Universal Robots PolyScope program: TgtProg.urp

Program TgtProg (createdIn=3.0.0 lastSavedIn=3.0.0 directory=/programs installation=default)
Robot Program (runOnlyOnce=true motionType=MoveJ speed=1.047198 acceleration=1.396263 useActiveTCP=false)
  'Program generated by RoboDK v6.0.7 for UR10 on XX/XX/XXXX 18:00:00'
  'Using nominal kinematics.'
  Wait Sleep waitTime=0.01
  Wait Sleep waitTime=0.01
  Wait Sleep waitTime=0.01
  Wait Sleep waitTime=0.01
  Wait Sleep waitTime=0.01
  Wait Sleep waitTime=0.01
